Staubli VAL3: copyPoint.pgx

public program copyPoint(string x_sKey, bool& x_bMark)
  local num l_nSize
  local num l_j
  local num l_i
begin
  resize(savedata:nMarkIndex,1,1)
  savedata:nMarkIndex=-1
  call getPointSize(x_sKey,l_nSize)
  l_j = 0
  for l_i = 0 to l_nSize-1
    if trajTemp:tTrajItem[x_sKey].pPointItem[l_i].bMarked
      l_j=l_j+1
      insert(savedata:nMarkIndex[l_j])
      savedata:nMarkIndex[l_j]=l_i


    endIf
  endFor
  x_bMark=false
end
